(* IEC 61131-3 sources: trust-platform/examples/rust_function_block/src/generated, 1 file *)

(* ---- rust_pous.st ---- *)
(* GENERATED by trust-runtime from rust/src/lib.rs - do not edit *)
{attribute 'rust'}
FUNCTION_BLOCK RAMP
VAR_INPUT
    EN : BOOL := TRUE;
    target : LREAL;
    rate : LREAL := 10.0;
END_VAR
VAR_OUTPUT
    out : LREAL;
    done : BOOL;
    ENO : BOOL;
END_VAR
END_FUNCTION_BLOCK
